Staubli VAL3: start.pgx

public program start()
begin
  call initArmInfo()
  call initWidget()
  call initDataBase()
  call mainCycle()
end
